// TIA Portal V19 export
VAR_GLOBAL   // PLC tag table "Conv"
   DI_Waffle_Insert AT %I8.0 : Bool;
   DI_Waffle_PickUpPosition AT %I8.1 : Bool;
   DI_Belt_Waffle_Conveyor AT %I8.4 : Bool;
END_VAR
